Staubli VAL3: modifyAll.pgx

public program modifyAll(string x_sKey, num x_nMoveType, num x_nParaSpeed, num x_nParaBlend, num x_nParaPercent, string x_sBlend, bool& x_bToSave, num x_nParaAcel)
  local num l_nSize
  local num l_i
begin
  call getPointSize(x_sKey,l_nSize)
  for l_i = 0 to l_nSize-1
    if trajTemp:tTrajItem[x_sKey].pPointItem[l_i].pParaItem.nMoveType==x_nMoveType
      // trajTemp:tTrajItem[x_sKey].pPointItem[l_i].pParaItem.nMoveType=x_nMoveType
      trajTemp:tTrajItem[x_sKey].pPointItem[l_i].pParaItem.mMdesc.vel=x_nParaSpeed
      trajTemp:tTrajItem[x_sKey].pPointItem[l_i].pParaItem.mMdesc.accel=x_nParaAcel
      trajTemp:tTrajItem[x_sKey].pPointItem[l_i].pParaItem.mMdesc.leave=x_nParaBlend
      trajTemp:tTrajItem[x_sKey].pPointItem[l_i].pParaItem.nPercentage=x_nParaPercent
      switch x_sBlend
        case "OFF"
          trajTemp:tTrajItem[x_sKey].pPointItem[l_i].pParaItem.mMdesc.blend=off
        break
        case "关节"
          trajTemp:tTrajItem[x_sKey].pPointItem[l_i].pParaItem.mMdesc.blend=joint
        break
        case "笛卡尔"
          trajTemp:tTrajItem[x_sKey].pPointItem[l_i].pParaItem.mMdesc.blend=Cartesian
        break
      endSwitch
    endIf
  endFor
  //trajTemp:libSave()
  //delay(0.5)
  logMsg("参数已修改")
  x_bToSave=true
end
